(* CODESYS project cognex_dm260.library
   DefaultNamespace: KOSTAL.AF2024.Drivers.Scanner.Cognex.DM260
   DocFormat: reStructuredText
   Description: Communication wit a Cognex Scanner Serie DM260
      Tested with real type DM262QX
   Author: Frank Dümpelmann
   Title: KOSTAL.AF2024.Drivers.Scanner.Cognex.DM260
   Version: 1.0.0.0
   Company: KOSTAL GmbH & Co.KG
   Placeholder: KOSTAL.AF2024.Drivers.Scanner.Cognex.DM260

Project tree, tasks and I/O mapping:
  libraries: KOSTAL.AF2024.Core.ListOf, 1.0.0.0 (KOSTAL GmbH & Co.KG); KOSTAL.AF2024.Core.Process, 1.0.0.0 (KOSTAL GmbH & Co.KG); KOSTAL.AF2024.Core.Settings, 1.0.0.0 (KOSTAL GmbH & Co.KG); KOSTAL.AF2024.Core.StringTools, 1.0.0.0 (KOSTAL GmbH & Co.KG); KOSTAL.AF2024.Core.System, 1.0.0.0 (KOSTAL GmbH & Co.KG); KOSTAL.AF2024.Drivers.Scanner.IScanner, 1.0.0.0 (KOSTAL GmbH & Co.KG); Tc2_Standard, 3.4.5.0 (Beckhoff Automation GmbH); Tc2_System, 3.6.4.0 (Beckhoff Automation GmbH); Tc2_TcpIp, 3.3.10.0 (Beckhoff Automation GmbH)
  Device/
    DUT/
      data type E_Command
      data type E_THIS
      data type T_SetupNumber
    POE/
      function block FB_Scanner [ST]: FB_init, _a0_stepFail, _a0_stepInit, _a1_Finish, _a1_Idle, _a2_Connect, _a2_Receive, _a2_Send, _a3_DisableSetup, _a3_EnableSetup, _a3_SelectSetup, _devices, _getCommand, _splitString, _timeOutOccured, _FBmain, ClearCodes, CodeGet, Ex_DisableSetup, Ex_EnableSetup, Ex_Scan, NativeStringGet, IP, Port, ExecutedSocketState, NumberOfBarcodes, serverAmsNetId, State, FBmain
      interface I_Scanner: Ex_DisableSetup, Ex_EnableSetup, ExecutedSocketState
  Project Information/
    function F_GetCompany [ST]
    function F_GetTitle [ST]
    function F_GetVersion [ST]
  Version/
    global variables Global_Version
*)

// Device/DUT/E_Command
{attribute 'qualified_only'}
{attribute 'strict'}
TYPE E_Command :
(
	TriggerOn := 0,
	TriggerOff,
	//UseSetupOn, do not use - setup will only hide - not disabled!
	//UseSetupOff, do not use - setup will only hide - not disabled!
	SelectSetup,
	EnableSetup,
	DisableSetup
);
END_TYPE

// Device/DUT/E_THIS
{attribute 'qualified_only'}
{attribute 'strict'}
TYPE E_THIS :
(
	Idle := 0,
	Scan,
	EnableSetup,
	DisableSetup
);
END_TYPE

// Device/DUT/T_SetupNumber

TYPE T_SetupNumber : UINT(0..15);END_TYPE

// Version/Global_Version
{attribute 'TcGenerated'}
{attribute 'no-analysis'}
{attribute 'linkalways'}
// This function has been automatically generated from the project information.
VAR_GLOBAL CONSTANT
	{attribute 'const_non_replaced'}
	stLibVersion_KOSTAL_AF2024_Drivers_Scanner_Cognex_DM260 : ST_LibVersion := (iMajor := 1, iMinor := 0, iBuild := 0, iRevision := 0, nFlags := 0, sVersion := '1.0.0.0');
END_VAR

// Device/POE/FB_Scanner
{info 'The Beckhoff Library >TF6310-TCP-IP.exe< is needed'}
(*

:Author: Frank Dümpelmann <f.duempelmann@kostal.com>, Martin Hundt <m.hundt@kostal.com>
:Date: 2019-01-07

Function
========
| Extension of FB_Reader to connect to a barcode reader via TCP/IP
| Tested with Keyence SR 750 

Usage notes
===============
| Asyncronous function block: FBmain() method must be called cyclicly
| The Beckhoff Library >TF6310-TCP-IP.exe< is needed

Methods and Properties
======================
| See bottom of this document for a detailed description of each method or property
| Methods starting with an underline(_) are internally used and can be ignored by the user

| Usage sample: ..\Device\Scanner\scannerBestPractice
| Usage Keyence Template ..\Device\Scanner\Keyence_SR\Keyence SR-750.ptc .. \Keyence SR-1000.ptc

*)
FUNCTION_BLOCK PUBLIC FB_Scanner IMPLEMENTS I_Scanner
VAR CONSTANT
		_PortDefault	: UDINT:= 23;
		_MaxSetup			: UDINT:= 15;
END_VAR
VAR

	_serverAmsNetId	: Tc2_System.T_AmsNetID:= '';
	_IP			: Tc2_System.T_IPv4Addr;
	_Port		: UDINT:= _PortDefault;

	_socket								: Tc2_TcpIp.FB_ClientServerConnection;
	_executedSocketState	:	Tc2_TcpIp.E_SocketConnectionState;
	
	_send						: Tc2_TcpIp.FB_SocketSend;
	_receive				: Tc2_TcpIp.FB_SocketReceive;

	_receivedPartly	: KOSTAL_AF2024_Core_Settings.T_MaxString_UTF8;
	//_receiveAck			: KOSTAL_AF2024_Core_Settings.T_MaxString_UTF8;


	_Command	: KOSTAL_AF2024_Core_Settings.T_MaxString_UTF8:= '||0:000>TRIGGER ON$0D$0A';	//default
	_STX									: STRING(1):= '$02';	//default	'$02';
	_ETX									: STRING(1):= '$03';	//default	'$03';
	_intermediateLimiter	: STRING(1):= '$04';

	_timeOut			: TIME	:= T#5S;	//default T#5S
	_timeOutTimer	: TON;	//TON

	
	_receivedString	: KOSTAL_AF2024_Core_Settings.T_MaxString_UTF8;
	_split					: KOSTAL_AF2024_Core_StringTools.FB_Split_UTF8;
	_barcodes				: KOSTAL_AF2024_Core_ListOf.FB_ListOfString_UTF8;
	
	_Step			: KOSTAL_AF2024_Core_Process.FB_processStep;
	_SubStep	: KOSTAL_AF2024_Core_Process.FB_processStep;
	_Init			: BOOL:= TRUE;

	_state		:	KOSTAL_AF2024_Core_Process.T_plcState;

	//_MaxAvailableSetupIndex	: T_SetupNumber:= 0;
	_SetupNumber						: T_SetupNumber:= 0;
	//_SelectedSetupNumber		: T_SetupNumber:= 0;
	//_PrepareSetupNumber		: T_SetupNumber:= 0;
	
	_THIS_CALLED			: E_THIS;
	_THIS_IN_PROCESS	: E_THIS;
	
	//_IndexCounter		: T_SetupNumber;
	//_LoopHeader			: INT;


END_VAR

VAR CONSTANT
	
	_SETUP_MAX_INDEX	: T_SetupNumber:= 15;
	
	_ADDRESS_READY					: INT:= 0;	
	_ADDRESS_ENABLE_SETUP		: INT:= 100;	
	_ADDRESS_DISABLE_SETUP	: INT:= 200;	
END_VAR

METHOD FB_init : BOOL
VAR_INPUT
	bInitRetains : BOOL; // if TRUE, the retain variables are initialized (warm start / cold start)
	bInCopyCode : BOOL;  // if TRUE, the instance afterwards gets moved into the copy code (online change)
	ServerAmsNetId	: Tc2_System.T_AmsNetID;
	Scanner_IP				: Tc2_System.T_IPv4Addr;
	Scanner_Port			: UDINT;
END_VAR

IF ServerAmsNetId <> ''	THEN	_serverAmsNetId:= serverAmsNetId;	END_IF
IF Scanner_IP <> ''			THEN	_IP:= Scanner_IP;									END_IF
IF Scanner_Port	<> 0		THEN	_Port:= Scanner_Port;							END_IF
END_METHOD

METHOD PROTECTED _a0_stepFail
VAR_INPUT
END_VAR

	_state.clear();
	_state.description:= Tc2_Standard.WCONCAT("Step does not exist: ", INT_TO_WSTRING(_step.actual));
	_state.fail		:= TRUE;
	_state.finish	:= TRUE;
END_METHOD

METHOD PUBLIC _a0_stepInit
VAR_INPUT
END_VAR

//Overwrite base method

IF _Init THEN

	_step.init();
	_Init:= FALSE;	

	_socket.bEnable		:= FALSE;
	_send.bExecute		:= FALSE;
	_receive.bExecute	:= FALSE;

	_timeOutTimer.IN:= FALSE;

ELSIF _THIS_CALLED <> _THIS_IN_PROCESS AND _step.actual > 0 THEN 

	_step.init();

	_socket.bEnable		:= FALSE;
	_send.bExecute		:= FALSE;
	_receive.bExecute	:= FALSE;

	_timeOutTimer.IN:= FALSE;

END_IF
END_METHOD

METHOD PROTECTED _a1_Finish
VAR_INPUT
END_VAR

IF _step.toggle THEN

	_timeOutTimer.IN:= FALSE;

	_socket.bEnable		:= FALSE;
	_send.bExecute		:= FALSE;
	_receive.bExecute	:= FALSE;

END_IF

_state.clear();
_state.finish	:= TRUE;
_state.pass		:= TRUE;
END_METHOD

METHOD PROTECTED _a1_Idle
VAR_INPUT
END_VAR

_state.clear();

_THIS_IN_PROCESS:= E_THIS.Idle;


IF _step.toggle THEN

	_socket(bEnable		:= FALSE);
	_send(bExecute		:= FALSE);
	_receive(bExecute	:= FALSE);

	_timeOutTimer(IN:= FALSE);

	_state.busy:= TRUE;

	
ELSIF 	_socket.bBusy THEN

	_state.busy:= TRUE;
	_state.description:= "socket is busy, please wait...";
	
ELSIF _send.bBusy THEN

	_state.busy:= TRUE;
	_state.description:= "send is busy, please wait...";

	
ELSIF _receive.bBusy THEN

	_state.busy:= TRUE;
	_state.description:= "receive is busy, please wait...";

ELSIF _THIS_CALLED = E_THIS.Idle THEN

	_state.ready:= TRUE;

	
ELSIF _THIS_CALLED = E_THIS.Scan THEN

	_THIS_IN_PROCESS:= _THIS_CALLED;

	_state.busy:= TRUE;

	_receivedString:= '';
	_receivedPartly:= '';
	
	_split.clear();
	_barcodes.clear();
	
	_timeOutTimer.IN:= TRUE;
	
	_state.clear();
	_state.busy:= TRUE;

	_Command	:= _getCommand(E_Command.TriggerOn, 0);

	_step.INC();
	
	
ELSIF _THIS_CALLED = E_THIS.EnableSetup THEN

	_THIS_IN_PROCESS:= _THIS_CALLED;

	IF _SetupNumber > _MaxSetup THEN
		
		_state.description:= "Number of setup is out of range (0..15)";
		_state.fail:= TRUE;
		_state.finish:= TRUE;

	ELSE

		_state.busy:= TRUE;
	
		_timeOutTimer.IN:= TRUE;
		
		_state.clear();
		_state.busy:= TRUE;

		_step.set(_ADDRESS_ENABLE_SETUP);
		
	END_IF

	
ELSIF _THIS_CALLED = E_THIS.DisableSetup THEN

	_THIS_IN_PROCESS:= _THIS_CALLED;

	IF _SetupNumber > _MaxSetup THEN
		
		_state.description:= "Number of setup is out of range (0..15)";
		_state.fail:= TRUE;
		_state.finish:= TRUE;

	ELSE

		_state.busy:= TRUE;
	
		_timeOutTimer.IN:= TRUE;
		
		_state.clear();
		_state.busy:= TRUE;

		_step.set(_ADDRESS_DISABLE_SETUP);
		
	END_IF

ELSE

	_state.clear();
	_state.ready:= TRUE;
		
END_IF
END_METHOD

METHOD PROTECTED _a2_Connect
VAR
	_c	: KOSTAL_AF2024_Core_StringTools.FB_Concat;
END_VAR

IF _step.toggle THEN
	_state.clear();
	_state.busy:= TRUE;
	_subStep.init();
END_IF


IF _timeOutTimer.Q THEN

	_timeOutOccured();

ELSE

	_subStep.Header();
	
	CASE _subStep.actual OF
		0:	_socket.bEnable:= FALSE;	_subStep.INC();
		1:	_socket.bEnable:= TRUE;		_subStep.INC();

		2:	IF _socket.bBusy THEN
					_state.busy	:= TRUE;
					_state.description:= "Scanner is busy(connect); wait ...";
				ELSE
					_subStep.INC();
				END_IF

		3:	IF _socket.bError THEN
					_state.clear();
					_state.description:= Tc2_Standard.WCONCAT("Error during socket open. Errorcode>", UDINT_TO_WSTRING(_socket.nErrId));
					_state.fail	:= TRUE;
					_state.finish:= TRUE;	
					_timeOutTimer.IN:= FALSE;
				ELSIF _socket.hSocket.handle = 0 THEN
					_state.clear();
					_state.description:= "no Handle from socket";
					_state.fail	:= TRUE;
					_state.finish:= TRUE;
					_timeOutTimer.IN:= FALSE;
				ELSE
					_step.INC();
				END_IF
		
	ELSE
	
		_timeOutTimer.IN:= FALSE;
		_state.clear();
		_state.fail	:= TRUE;
		_state.finish:= TRUE;
		_c.clear();
		_c.addContent("connect Step ");
		_c.addContent(INT_TO_WSTRING(_subStep.actual));
		_c.addContent(" does not exist");
		_state.description:= _c.getResult();
		_c.clear();
	
	END_CASE

END_IF
END_METHOD

METHOD PROTECTED _a2_Receive
VAR
	_c	: KOSTAL_AF2024_Core_StringTools.FB_Concat;
END_VAR

IF _step.toggle THEN

	_state.clear();
	_state.busy:= TRUE;

	_subStep.init();

	_receivedString:= '';
	_receivedPartly:= '';

	_split.clear();
	_barcodes.clear();

END_IF



IF _timeOutTimer.Q THEN

	_timeOutOccured();

ELSE
	
	_subStep.Header();

	CASE _subStep.actual OF
		0:	_receive.bExecute:= FALSE;	_receivedPartly:= '';	_subStep.INC();
		1:	_receive.bExecute:= TRUE;		_subStep.INC();

		2:	IF _receive.bBusy THEN
					_state.busy	:= TRUE;
					_state.description:= "Scanner is busy(receive); wait ...";
				ELSE
					_subStep.INC();
				END_IF

		3:	IF _receive.bError THEN
					_state.clear();
					_state.description:= Tc2_Standard.WCONCAT("Error during receive. Errorcode>", UDINT_TO_WSTRING(_receive.nErrId));
					_state.fail	:= TRUE;
					_state.finish:= TRUE;	
					_timeOutTimer.IN:= FALSE;
				ELSE
					_subStep.INC();
				END_IF
		
		4:	IF	_receive.nRecBytes <> 0 THEN 

					_receivedString:= Tc2_Standard.CONCAT(STR1:= _receivedString, STR2:=  Tc2_Standard.LEFT(STR:= _receivedPartly, SIZE:= UDINT_TO_INT(_receive.nRecBytes)));
					_receivedPartly:= '';
					_splitString();

					_subStep.SET(0);

				ELSIF (_barcodes.NumberOfLines < 1) THEN 

					_subStep.SET(0);

				ELSE
					
					_state.clear();
					_state.busy:= TRUE;
					_state.pass:= TRUE;
					_timeOutTimer.IN:= FALSE;
					_step.INC();

				END_IF
								
	ELSE
	
		_timeOutTimer.IN:= FALSE;
		_state.clear();
		_state.fail	:= TRUE;
		_state.finish:= TRUE;
		_c.clear();
		_c.addContent("send Step ");
		_c.addContent(INT_TO_WSTRING(_subStep.actual));
		_c.addContent(" does not exist");
		_state.description:= _c.getResult();
		_c.clear();
	
	END_CASE

END_IF
END_METHOD

METHOD PROTECTED _a2_Send
VAR
	_c	: KOSTAL_AF2024_Core_StringTools.FB_Concat;
END_VAR

IF _step.toggle THEN
	_state.clear();
	_state.busy:= TRUE;
	_subStep.init();
END_IF


IF _timeOutTimer.Q THEN

	_timeOutOccured();

ELSE
	
	_subStep.Header();

	CASE _subStep.actual OF
		0:	_send.bExecute:= FALSE;	_subStep.INC();
		1:	_send.bExecute:= TRUE;		_subStep.INC();

		2:	IF _send.bBusy THEN
					_state.busy	:= TRUE;
					_state.description:= "Scanner is busy(send); wait ...";
				ELSE
					_subStep.INC();
				END_IF

		3:	IF _send.bError THEN
					_state.clear();
					_state.description:= Tc2_Standard.WCONCAT("Error during send. Errorcode>", UDINT_TO_WSTRING(_send.nErrId));
					_state.fail	:= TRUE;
					_state.finish:= TRUE;	
					_timeOutTimer.IN:= FALSE;
				ELSE
					_step.INC();
				END_IF
		
	ELSE
	
		_state.clear();
		_state.fail	:= TRUE;
		_state.finish:= TRUE;
		_c.clear();
		_c.addContent("send Step ");
		_c.addContent(INT_TO_WSTRING(_subStep.actual));
		_c.addContent(" does not exist");
		_state.description:= _c.getResult();
		_c.clear();
	
	END_CASE

END_IF
END_METHOD

METHOD PROTECTED _a3_DisableSetup
VAR_INPUT
END_VAR


_Command	:= _getCommand(E_Command.DisableSetup, _SetupNumber);

_Step.INC();
END_METHOD

METHOD PROTECTED _a3_EnableSetup
VAR_INPUT
END_VAR
	
_Command	:= _getCommand(E_Command.EnableSetup, _SetupNumber);

_Step.INC();
END_METHOD

METHOD PROTECTED _a3_SelectSetup
VAR_INPUT
END_VAR


_Command	:= _getCommand(E_Command.SelectSetup, _SetupNumber);

_Step.INC();
END_METHOD

METHOD PROTECTED _devices
VAR_INPUT
END_VAR


_timeOutTimer(IN:= , PT:= _timeOut, Q=> , ET=> );

_socket
	(
		sSrvNetID	:= _serverAmsNetId, 
		nMode			:= Tc2_TcpIp.CONNECT_MODE_ENABLEDBG, 

		sRemoteHost	:= _IP, 
		nRemotePort	:= _Port, 

		bEnable			:= , 
		tReconnect	:= _timeOut, 

		bBusy		=> , 
		bError	=> , 
		nErrId	=> , 
		hSocket	=> , 
		eState	=> 
	);
	
IF _socket.bEnable THEN	_executedSocketState:= _socket.eState;	END_IF
	
_send
	(
		sSrvNetId	:= _serverAmsNetId, 
		hSocket		:= _socket.hSocket, 
		cbLen			:= SIZEOF(_Command), 
		pSrc			:= ADR(_Command), 
		bExecute	:= , 
		tTimeout	:= _timeOut, 

		bBusy			=> , 
		bError		=> , 
		nErrId		=> 
	);
	
	
	_receive
	(
		sSrvNetId	:= _serverAmsNetId, 
		hSocket		:= _socket.hSocket, 

		cbLen:= SIZEOF(_receivedPartly) - 1, 
		pDest:= ADR(_receivedPartly), 

		bExecute:= , 
		tTimeout:= _timeOut, 

		bBusy			=> , 
		bError		=> , 
		nErrId		=> , 
		nRecBytes	=> 
	);
END_METHOD

METHOD PROTECTED _getCommand : KOSTAL_AF2024_Core_Settings.T_MaxString_UTF8

VAR_INPUT
	ID				: E_Command;
	Parameter : UINT;
END_VAR
VAR
	_c	: KOSTAL_AF2024_Core_StringTools.FB_Concat_UTF8;
END_VAR

CASE ID OF
	E_Command.TriggerOn		: _getCommand:= '||0:000>TRIGGER ON$0D$0A';
	
	E_Command.TriggerOff	: _getCommand:= '||0:000>TRIGGER OFF$0D$0A';

	(* do not use - setup will only hide - not disabled!
		=====================================================================
	E_Command.UseSetupOn		: _c.clear();
														_c.addContent('||0:000>SETUP.USE ');
														_c.addContent(UINT_TO_STRING(Parameter));
														_c.addContent(' ON');
														_c.addContent('$0D$0A');
														_getCommand:= _c.getResult();
														_c.clear();
														
	E_Command.UseSetupOff		: _c.clear();
														_c.addContent('||0:000>SETUP.USE ');
														_c.addContent(UINT_TO_STRING(Parameter));
														_c.addContent(' OFF');
														_c.addContent('$0D$0A');
														_getCommand:= _c.getResult();
														_c.clear();
		=====================================================================
*)
														
	E_Command.SelectSetup	: _c.clear();
													_c.addContent('||0:000>SET SETUP.PROG-TARGET ');
													_c.addContent(UINT_TO_STRING(Parameter));
													_c.addContent('$0D$0A');
													_getCommand:= _c.getResult();
													_c.clear();
	
	E_Command.EnableSetup	: _c.clear();
													_c.addContent('||0:000>SET SETUP.ENABLE ');
													_c.addContent('ON');
													_c.addContent('$0D$0A');
													_getCommand:= _c.getResult();
													_c.clear();
													
	E_Command.DisableSetup	: _c.clear();
														_c.addContent('||0:000>SET SETUP.ENABLE ');
														_c.addContent('OFF');
														_c.addContent('$0D$0A');
														_getCommand:= _c.getResult();
														_c.clear();

END_CASE
END_METHOD

(*
| split received string depends of STX ETX
*)
METHOD PROTECTED _splitString  : BOOL

VAR
	_udi: UDINT;
	_element: KOSTAL_AF2024_Core_Settings.T_MaxString_UTF8;
	_stxPos: INT;
	_code: KOSTAL_AF2024_Core_Settings.T_MaxString_UTF8;
END_VAR
_barcodes.clear();

IF _receivedString = '' THEN
	
	;	// no splitting possible

	
// if EXT is defined
// ============================================================================
ELSIF _ETX <> '' THEN

	_split.clear();
	_split.Delimiter:= _ETX;
	_split.split(_receivedString);

	// if additional STX is defined then select
	IF _STX <> '' THEN

		FOR _udi:= 1 TO _split.Results.NumberOfLines DO
			
			_element:= _split.Results.line_GET(_udi);
			_stxPos:= Tc2_Standard.FIND(STR1:= _element, STR2:= _STX);

			IF _stxPos > 0 THEN
				_barcodes.addLine(newLine:= Tc2_Standard.RIGHT(STR:= _element, SIZE:= Tc2_Standard.LEN( STR:= _element) - _stxPos ));
			END_IF
		END_FOR
	
	// no STX defined
	ELSE

		FOR _udi:= 1 TO _split.Results.NumberOfLines DO
			_barcodes.addLine(newLine:= _split.Results.line_GET(_udi));
		END_FOR
	
	END_IF

	
// if only STX is defined
// ============================================================================
ELSIF _STX <> '' THEN
	
	_split.clear();
	_split.Delimiter:= _STX;
	_split.split(_receivedString);

	FOR _udi:= 1 TO _split.Results.NumberOfLines DO
		_barcodes.addLine(newLine:= _split.Results.line_GET(_udi));
	END_FOR

// neither STX or ETX is defined then no splitting possible
// ============================================================================
ELSE

	_barcodes.addLine(newLine:= _receivedString);

END_IF

_splitString:= _barcodes.NumberOfLines > 0;

IF _barcodes.NumberOfLines = 1 THEN

	_code:= _barcodes.line_GET(1);

	_split.clear();
	_split.Delimiter:= _intermediateLimiter;
	_split.split(_code);

	_barcodes.removeLine(1);

	FOR _udi:= 1 TO _split.Results.NumberOfLines DO
		_barcodes.addLine(_split.Results.line_GET(_udi));
	END_FOR


END_IF
END_METHOD

METHOD PROTECTED _timeOutOccured
VAR_INPUT
END_VAR


_socket.bEnable		:= FALSE;
_send.bExecute		:= FALSE;
_receive.bExecute	:= FALSE;

_state.busy:= FALSE;
_state.description:= "Timeout";
_state.fail:= TRUE;
_state.finish:= TRUE;
END_METHOD

(*
Decription
==========
*)
METHOD PROTECTED _FBmain


_a0_stepInit();

_step.Header();

CASE _step.actual OF

	0:	_a1_Idle();
	
	1:	_a2_Connect();
	2:	_a2_Send();
	3:	_a2_Receive();
	4:	_a1_Finish();

(*
	_ADDRESS_SET_MAX_INDEX:	_IndexCounter:= 1;	 _step.INC();
	101:	_a2_Connect();
	102:	_a4_LoopHeader_MaxIndex(); 
	103:	_a2_Send();
	104:	_a4_LoopBottom();

*)
	_ADDRESS_ENABLE_SETUP:	_step.INC();
	101:	_a2_Connect();
	102:	_a3_SelectSetup();
	103:	_a2_Send();
	104:	_a3_EnableSetup();
	105:	_a2_Send();
	106:	_a1_Finish();

	_ADDRESS_DISABLE_SETUP:	_step.INC();
	201:	_a2_Connect();
	202:	_a3_SelectSetup();
	203:	_a2_Send();
	204:	_a3_DisableSetup();
	205:	_a2_Send();
	206:	_a1_Finish();

ELSE	_a0_stepFail();	

END_CASE
	
	

_devices();
END_METHOD

METHOD PUBLIC ClearCodes

_barcodes.clear();
_receivedString:= '';
END_METHOD

METHOD PUBLIC CodeGet : KOSTAL_AF2024_Core_Settings.T_MaxString_UTF8
VAR_INPUT
	number	: UINT;
END_VAR

IF (number = 0) OR (number > _barcodes.NumberOfLines) THEN
	CodeGet:= '';
ELSE
	CodeGet:= _barcodes.line_GET(number);
END_IF
END_METHOD

METHOD Ex_DisableSetup : BOOL

VAR_INPUT
	SetupNumber	: T_SetupNumber;
END_VAR
IF _THIS_CALLED = E_THIS.Idle THEN

	_THIS_CALLED:= E_THIS.DisableSetup;

	_SetupNumber:= SetupNumber;

	_FBmain();

	Ex_DisableSetup:= _THIS_CALLED = _THIS_IN_PROCESS;
	
ELSE
	
	Ex_DisableSetup:= FALSE;
 
END_IF
END_METHOD

METHOD Ex_EnableSetup : BOOL

VAR_INPUT
	SetupNumber	: T_SetupNumber;
END_VAR
IF _THIS_CALLED = E_THIS.Idle THEN

	_THIS_CALLED:= E_THIS.EnableSetup;

	_SetupNumber:= SetupNumber;

	_FBmain();

	Ex_EnableSetup:= _THIS_CALLED = _THIS_IN_PROCESS;
	
ELSE
	
	Ex_EnableSetup:= FALSE;
 
END_IF
END_METHOD

METHOD Ex_Scan : BOOL
IF _THIS_CALLED = E_THIS.Idle THEN

	_THIS_CALLED:= E_THIS.Scan;

	_FBmain();

	Ex_Scan:= _THIS_CALLED = _THIS_IN_PROCESS;

ELSE

	Ex_Scan:= FALSE;
	
END_IF
END_METHOD

METHOD PUBLIC NativeStringGet : KOSTAL_AF2024_Core_Settings.T_MaxString_UTF8
VAR_INPUT
END_VAR

NativeStringGet:= _receivedString;
END_METHOD

(*
Description
===========
| IP address of the barcode reader
*)
PROPERTY PUBLIC IP : STRING
GET


IP:= _IP;
END_GET
SET

_IP:= IP;
END_SET
END_PROPERTY

(*
Description
===========
| TCP/IP port of the barcode reader
*)
PROPERTY PUBLIC Port : UDINT
GET


Port:= _Port;
END_GET
SET

IF Port = UDINT#0 THEN	_Port:= _PortDefault;
ELSE										_Port:= Port;
END_IF
END_SET
END_PROPERTY

(*
Description
===========
| State of the TCP/IP connection
*)
PROPERTY PUBLIC ExecutedSocketState : E_SocketConnectionState
GET

ExecutedSocketState:= _executedSocketState;
END_GET
END_PROPERTY

PROPERTY PUBLIC NumberOfBarcodes : UDINT
GET

NumberOfBarcodes:= _barcodes.NumberOfLines;
END_GET
END_PROPERTY

(*
Description
===========
| AmsNetId of the system running the Beckhoff TCP/IP server
| default: ''=local system
*)
PROPERTY PUBLIC serverAmsNetId : STRING
GET

serverAmsNetId:= _serverAmsNetId;
END_GET
SET

_serverAmsNetId:= serverAmsNetId;
END_SET
END_PROPERTY

PROPERTY PUBLIC State : KOSTAL_AF2024_Core_Process.I_T_plcState
GET

State:= _state;
END_GET
END_PROPERTY

(*
Decription
==========
| To be called cyclicly, e.g. in DeviceDefine
*)
METHOD PUBLIC FBmain
VAR_INPUT
END_VAR

IF _THIS_CALLED = E_THIS.Idle THEN
	_FBmain();
END_IF

_THIS_CALLED:= E_THIS.Idle;
END_METHOD

END_FUNCTION_BLOCK

// Device/POE/I_Scanner
INTERFACE I_Scanner EXTENDS KOSTAL_AF2024_Drivers_Scanner_IScanner.I_Scanner

METHOD Ex_DisableSetup : BOOL

VAR_INPUT
	SetupNumber	: T_SetupNumber;
END_VAR
END_METHOD

METHOD Ex_EnableSetup : BOOL
VAR_INPUT
	SetupNumber	: T_SetupNumber;
END_VAR
END_METHOD

(*
Description
===========
| State of the TCP/IP connection
*)
PROPERTY PUBLIC ExecutedSocketState : E_SocketConnectionState
GET
END_GET
END_PROPERTY

END_INTERFACE

// Project Information/F_GetCompany
// This function has been automatically generated from the project information.
{attribute 'signature_flag' := '1073741824'}
{attribute 'TcGenerated'}
{attribute 'no-analysis'}
FUNCTION F_GetCompany : WSTRING
VAR_INPUT
	
END_VAR

F_GetCompany := "KOSTAL GmbH & Co.KG";

END_FUNCTION

// Project Information/F_GetTitle
// This function has been automatically generated from the project information.
{attribute 'signature_flag' := '1073741824'}
{attribute 'TcGenerated'}
{attribute 'no-analysis'}
FUNCTION F_GetTitle : WSTRING
VAR_INPUT
	
END_VAR

F_GetTitle := "KOSTAL.AF2024.Drivers.Scanner.Cognex.DM260";

END_FUNCTION

// Project Information/F_GetVersion
// This function has been automatically generated from the project information.
{attribute 'signature_flag' := '1073741824'}
{attribute 'TcGenerated'}
{attribute 'no-analysis'}
FUNCTION F_GetVersion : ST_LibVersion
VAR_INPUT
	
END_VAR

F_GetVersion.iMajor := 1;
F_GetVersion.iMinor := 0;
F_GetVersion.iBuild := 0;
F_GetVersion.iRevision := 0;
F_GetVersion.sVersion := '1.0.0.0';
F_GetVersion.nFlags := 0;

END_FUNCTION
